// TIA Portal V18 export
// export: Created 2026-11-25T00:00:00.0000000Z, ExportSetting WithDefaults
TagTable "Station"
  State : Int  (%DB{DB}.DBW0, Connection_PLC, 1 s)
  Verdict : Int  (%DB{DB}.DBW2, Connection_PLC, 1 s)
  NokCode : Int  (%DB{DB}.DBW4, Connection_PLC, 1 s)
  FaultCode : Int  (%DB{DB}.DBW6, Connection_PLC, 1 s)
  CntConsecNok : Int  (%DB{DB}.DBW8, Connection_PLC, 1 s)
  Locked : Bool  (%DB{DB}.DBX10.0, Connection_PLC, 1 s)
  RigCheck : Bool  (%DB{DB}.DBX10.1, Connection_PLC, 1 s)
  CallOperator : Bool  (%DB{DB}.DBX10.2, Connection_PLC, 1 s)
  PartPresent : Bool  (%DB{DB}.DBX10.3, Connection_PLC, 1 s)
  TCycle : Real  (%DB{DB}.DBD12, Connection_PLC, 1 s)
  CntTotal : DInt  (%DB{DB}.DBD16, Connection_PLC, 1 s)
  CntOk : DInt  (%DB{DB}.DBD20, Connection_PLC, 1 s)
  CntNok : DInt  (%DB{DB}.DBD24, Connection_PLC, 1 s)
  CntRejectConfirmed : DInt  (%DB{DB}.DBD28, Connection_PLC, 1 s)
  FpG1 : Real  (%DB{DB}.DBD32, Connection_PLC, 1 s)
  FrG1 : Real  (%DB{DB}.DBD36, Connection_PLC, 1 s)
  FMean : Real  (%DB{DB}.DBD40, Connection_PLC, 1 s)
  FHyst : Real  (%DB{DB}.DBD44, Connection_PLC, 1 s)
  FpG2 : Real  (%DB{DB}.DBD48, Connection_PLC, 1 s)
  FPeak : Real  (%DB{DB}.DBD52, Connection_PLC, 1 s)
  XPeak : Real  (%DB{DB}.DBD56, Connection_PLC, 1 s)
  FStep : Real  (%DB{DB}.DBD60, Connection_PLC, 1 s)
  XStop : Real  (%DB{DB}.DBD64, Connection_PLC, 1 s)
  MeanLo : Real  (%DB{DB}.DBD68, Connection_PLC, 1 s)
  MeanHi : Real  (%DB{DB}.DBD72, Connection_PLC, 1 s)
  HystLo : Real  (%DB{DB}.DBD76, Connection_PLC, 1 s)
  HystHi : Real  (%DB{DB}.DBD80, Connection_PLC, 1 s)
  G2Lo : Real  (%DB{DB}.DBD84, Connection_PLC, 1 s)
  G2Hi : Real  (%DB{DB}.DBD88, Connection_PLC, 1 s)
  PeakFLo : Real  (%DB{DB}.DBD92, Connection_PLC, 1 s)
  PeakFHi : Real  (%DB{DB}.DBD96, Connection_PLC, 1 s)
  PeakXMin : Real  (%DB{DB}.DBD100, Connection_PLC, 1 s)
  PeakXMax : Real  (%DB{DB}.DBD104, Connection_PLC, 1 s)
  StepLo : Real  (%DB{DB}.DBD108, Connection_PLC, 1 s)
  StopXLo : Real  (%DB{DB}.DBD112, Connection_PLC, 1 s)
  StopXHi : Real  (%DB{DB}.DBD116, Connection_PLC, 1 s)
